Universal Robots URScript: T002_codellama_34b_adversarial_A8.1_rep1.urscript

def linear_weld_path():
    # Move to home position
    movej(p[300.0, 0.0, 0.0, 0.0, 0.0, 0.0], v=300.0)

    # Approach above weld start
    movel(p[250.0, 0.0, 0.0, 0.0, 0.0, 0.0], v=250.0)

    # Descend
